FUNCTION_BLOCK DlPgnSend (* Send a PGN once without an installed Tx PGN *)
  (* Standard: 61499-2; Description: Calls iso_DlPgnSend() of the CCI ISOBUS driver (data link layer). \n 0..8 bytes are sent as single frame, 9..1785 bytes with TP (NMEA 2000 PGNs with Fast Packet). \n More than 1785 bytes (ETP) are refused with s16Status E_RANGE, because the driver does not copy them. \n Sender is NmDestin.s16OwnCfHnd, receiver is NmDestin.s16Handle (HANDLE::GLOBAL for broadcast). \n Missing bytes (u16DaSize larger than Data) are sent as 0xFF. *)
  (* Version 1.0, 2026-11-17, Franz Höpfinger, initial API and implementation and/or initial documentation *)
  PACKAGE isobus::pgn::tx;
  IMPORT isobus::pgn::ISONETEVENT_T;
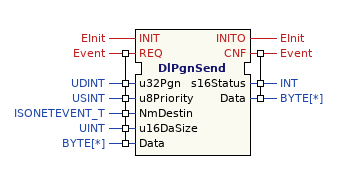
  EVENT_INPUT
    INIT : EInit; (* Service Initialization *)
    REQ WITH u32Pgn, u8Priority, NmDestin, u16DaSize, Data; (* Send the PGN once *)
  END_EVENT
  EVENT_OUTPUT
    INITO : EInit; (* Initialization Confirm *)
    CNF WITH s16Status, Data; (* Send started (see s16Status) *)
  END_EVENT
  VAR_INPUT
    u32Pgn : UDINT; (* PGN - Range: 0 - 0x3FFFF *)
    u8Priority : USINT := 6; (* Priority (0..7) 0=highest *)
    NmDestin : isobus::pgn::ISONETEVENT_T; (* Sender (s16OwnCfHnd) and receiver (s16Handle) *)
    u16DaSize : UINT; (* Number of data bytes to send (0..1785) *)
  END_VAR
  VAR_OUTPUT
    s16Status : INT; (* Return value of iso_DlPgnSend(): 0 = OK *)
  END_VAR
  VAR_IN_OUT
    Data : ARRAY [*] OF BYTE; (* data buffer *)
  END_VAR
END_FUNCTION_BLOCK
